Staubli VAL3: SmartTCP_CS9.pjx

--- SmartTCP_CS9.pjx ---
Parameters version=s8.10.5Cs9_BS2172 stackSize=20000 millimeterUnit=true
Program file=start.pgx
Program file=stop.pgx
Program file=V20201012.pgx
Data file=SmartTCP_CS9.dtx
Library alias=tx2 path=./tx2/tx2.pjx
Library alias=ts2 path=./ts2/ts2.pjx

--- SmartTCP_CS9.dtx ---


--- start.pgx ---
public program start()
  local string l_sArmType
  local string l_sSeries
begin
  //****************************************************************************************
  // +-----------------------------------------------------------------------------------+
  // !                                 Stäubli SmartTCP                                  !
  // !                                                                                   !
  // !                Copyright by  Stäubli(Hagnzhou) Mechatronic Co.,Ltd.               !
  // +-----------------------------------------------------------------------------------+
  // General description：  Stäubli TCP calibration application for TX2/TS2 robot
  // Developer:             ZhangHuaJun
  // Application version：  V1.2
  // Application Date:      February 24, 2020
  // Hardware required：    TX2/TS2-CS9-SP2 Robot
  // Software required：    Val3 s8.8.3+
  // VAL3 Addons：          Expansion
  // Fieldbus required:     None
  // VAL3 Options：         None
  // Included libraries：   None
  // Miscellaneous：        None
  //****************************************************************************************
  l_sArmType=getVersion("Arm Type")
  if l_sArmType!=""
    l_sSeries=left(l_sArmType,3)
    switch l_sSeries
      case "ts2"
        call ts2:start()
      break
      case "tx2"
        call tx2:start()
      break
    endSwitch
  endIf
end

--- stop.pgx ---
program stop()
begin
end

--- V20201012.pgx ---
program V20201012()
begin
  //Version: V1.2
  //Date: February 14, 2020
  //Editor: Zhang Huajun
  //  1.Improved real-time position display, can view joints and Cartesian coordinates
  //  2.Improve popup information display
  //  3.Corrected the error that the target point cannot be reached

  //Version: V1.3
  //Date: April 9, 2020
  //Editor: Zhang Huajun
  //  1.Reduce unnecessary binding
  //  2.Use CSS to keep Stäubli SP2 interface style
  //
  //
  //Version: V2.0
  //Date: August 20, 2020
  //Editor: Zhang Huajun
  //  1.Optimize HMI response by turning libsave() into a background task
  //  2.Optimize widgets binding
  //
  //
  //Version: V2.1
  //Date: October 12, 2020
  //Editor: Zhang Huajun
  //  1.Add 2 points to calculate TCP for 4-axis robot (only output X and Y)
end
